{region 'Documentation'}
(*!
<summary>Exercises the real UpdateStatus mapping and counts Prepare calls without resource actions.</summary>
*)
{endregion}
FUNCTION_BLOCK PreparationStatusProbe EXTENDS PreparationBase
VAR_INPUT
    DiagnosticState : E_State := E_State.Idle; //! Scripted diagnostic state projected by Prepare.
    ExecutionStatus : E_ExecutionStatus := E_ExecutionStatus.Idle; //! Scripted execution classification projected by Prepare.
    Ready : BOOL := TRUE; //! Scripted readiness projected by Prepare.
END_VAR
VAR
    FCallCount : UDINT;
END_VAR

SUPER^();

{region 'Documentation'}
(*!
<summary>Current CallCount observation.</summary>
*)
{endregion}
{attribute 'monitoring' := 'call'}
PROPERTY PUBLIC CallCount : UDINT //! Current CallCount observation.
GET // PUBLIC
CallCount := FCallCount;
END_GET
END_PROPERTY

{region 'Documentation'}
(*!
<summary>Calls the inherited status projector once, including when disabled.</summary>
*)
{endregion}
METHOD PROTECTED Prepare
FCallCount := FCallCount + 1;
UpdateStatus(State := DiagnosticState,
    ExecutionStatus := ExecutionStatus,
    Ready := Ready);
END_METHOD

END_FUNCTION_BLOCK

(* stored: Version 1.1.0.1
   POU PreparationStatusProbe: Id {651cff2e-d963-49f4-8693-1e0e50319d16}, SpecialFunc None
   Folder Internal: Id {3826a284-3aff-47b0-b279-06043bc7462c}
   Property CallCount: Id {4ea25e0f-8848-42ca-8846-7e49897fb3f7}
   Get Get: Id {dd8e9009-a703-4ddb-92f6-883627137434}
   Method Prepare: Id {af46e5dc-fbda-4963-bf25-1c1f75f38b39} *)
